(* IEC 61131-3 sources: PLC-Static-Analysis/modules/plc-rules/src/test/resources/PLCA-L020, 2 files *)

(* ---- compliant.st ---- *)
PROGRAM P_L020ok
VAR
    n : INT;
    m : INT;
    r : REAL;
    b : BOOL;
    c : BOOL;
    q : BOOL;
END_VAR
IF n > 10 THEN
    n := 0;
    q := TRUE;
ELSE
    n := 0;
    q := FALSE;
END_IF
IF n > 10 THEN
    q := TRUE;
    m := 0;
ELSIF n > 5 THEN
    q := FALSE;
    m := 0;
END_IF
IF n > 10 THEN
    q := TRUE;
    m := 0;
ELSE
    q := FALSE;
    m := 1;
END_IF
END_PROGRAM

(* ---- noncompliant.st ---- *)
PROGRAM P_L020
VAR
    n : INT;
    m : INT;
    r : REAL;
    b : BOOL;
    c : BOOL;
    q : BOOL;
END_VAR
IF n > 10 THEN
    q := TRUE;
    m := 0; // PLCA-L020
ELSE
    q := FALSE;
    m := 0;
END_IF
CASE n OF
    1: b := TRUE; // PLCA-L020
       q := TRUE;
    2: b := TRUE;
       q := FALSE;
ELSE
    b := TRUE;
END_CASE
END_PROGRAM
